(* IEC 61131-3 sources: llm-plc-st-eval/data/processed_definitivo/gemini-3.1-pro-preview/I5/zero_shot, 3 files *)

(* ---- ejec_1.st ---- *)
FUNCTION_BLOCK FB_Clasificadora
VAR_INPUT
    sensorPresencia : BOOL; // Sensor que detecta el paso de una pieza
    sensorAltura : BOOL;    // Sensor que detecta si la pieza es alta
END_VAR

VAR_OUTPUT
    banda : BOOL;           // Salida para activar la banda transportadora
    piston : BOOL;          // Salida para activar el pistón desviador
    nAltas : INT := 0;      // Contador de piezas altas
    nBajas : INT := 0;      // Contador de piezas bajas
END_VAR

VAR
    trigPresencia : R_TRIG; // Detector de flanco de subida para el sensor de presencia
    esperaPiston : BOOL;    // Marca de memoria para iniciar el retardo del pistón
    tonRetardo : TON;       // Temporizador de retardo (llegada al desviador)
    tpPiston : TP;          // Temporizador de pulso (duración de activación del pistón)
END_VAR

// 1. La banda funciona continuamente
banda := TRUE;

// 2. Detección del paso de una pieza (flanco de subida)
trigPresencia(CLK := sensorPresencia);

IF trigPresencia.Q THEN
    IF sensorAltura THEN
        // Es una pieza alta
        nAltas := nAltas + 1;
        esperaPiston := TRUE; // Se activa la bandera para iniciar el retardo
    ELSE
        // Es una pieza baja
        nBajas := nBajas + 1;
    END_IF;
END_IF;

// 3. Temporizador de retardo: espera 2 segundos a que la pieza llegue al pistón
tonRetardo(IN := esperaPiston, PT := T#2S);

// Al cumplirse los 2 segundos, se apaga la marca de espera
IF tonRetardo.Q THEN
    esperaPiston := FALSE;
END_IF;

// 4. Temporizador de pulso: activa el pistón durante 1 segundo
// Se dispara con el flanco de subida de tonRetardo.Q
tpPiston(IN := tonRetardo.Q, PT := T#1S);

// 5. Asignación de la salida física del pistón
piston := tpPiston.Q;

END_FUNCTION_BLOCK

(* ---- ejec_2.st ---- *)
FUNCTION_BLOCK FB_Clasificadora
VAR_INPUT
    sensorPresencia : BOOL; (* Detecta el paso de una pieza *)
    sensorAltura    : BOOL; (* Detecta si la pieza es alta *)
END_VAR
VAR_OUTPUT
    banda   : BOOL; (* Control de la banda transportadora *)
    piston  : BOOL; (* Control del pistón desviador *)
    nAltas  : INT;  (* Contador de piezas altas *)
    nBajas  : INT;  (* Contador de piezas bajas *)
END_VAR
VAR
    flancoPresencia : R_TRIG; (* Detector de flanco para contar solo una vez por pieza *)
    esperaPiston    : BOOL;   (* Marca para iniciar el retardo del pistón *)
    timerRetardo    : TON;    (* Temporizador para el tiempo de viaje (2s) *)
    timerPiston     : TP;     (* Temporizador para la duración del pistón (1s) *)
END_VAR

(* La banda está siempre activa *)
banda := TRUE;

(* Detectar el flanco de subida del sensor de presencia *)
flancoPresencia(CLK := sensorPresencia);

(* Lógica de clasificación y conteo al detectar una pieza *)
IF flancoPresencia.Q THEN
    IF sensorAltura THEN
        nAltas := nAltas + 1;
        esperaPiston := TRUE; (* Activa la bandera para iniciar el retardo *)
    ELSE
        nBajas := nBajas + 1;
    END_IF;
END_IF;

(* Temporizador TON: espera 2 segundos desde que se detecta la pieza alta *)
timerRetardo(IN := esperaPiston, PT := T#2S);

(* Cuando pasan los 2 segundos, se resetea la marca de espera *)
IF timerRetardo.Q THEN
    esperaPiston := FALSE;
END_IF;

(* Temporizador TP: genera un pulso de 1 segundo para el pistón *)
(* Se dispara exactamente cuando timerRetardo.Q se activa *)
timerPiston(IN := timerRetardo.Q, PT := T#1S);

(* Asignar la salida del temporizador al pistón *)
piston := timerPiston.Q;

END_FUNCTION_BLOCK

(* ---- ejec_3.st ---- *)
FUNCTION_BLOCK FB_Clasificadora
VAR_INPUT
    sensorPresencia : BOOL; (* Sensor que detecta el paso de una pieza *)
    sensorAltura : BOOL;    (* Sensor que detecta si la pieza es alta *)
END_VAR

VAR_OUTPUT
    banda : BOOL;           (* Salida para activar la banda transportadora *)
    piston : BOOL;          (* Salida para activar el pistón desviador *)
    nAltas : INT := 0;      (* Contador de piezas altas *)
    nBajas : INT := 0;      (* Contador de piezas bajas *)
END_VAR

VAR
    trigPresencia : R_TRIG; (* Detector de flanco de subida para la presencia *)
    tonRetardo : TON;       (* Temporizador para el retardo de 2 segundos *)
    tpPiston : TP;          (* Temporizador de pulso para el pistón de 1 segundo *)
    esperandoPiston : BOOL := FALSE; (* Memoria para el retardo del pistón *)
END_VAR

(* 1. La banda funciona continuamente *)
banda := TRUE;

(* 2. Detección de nueva pieza (flanco de subida) *)
trigPresencia(CLK := sensorPresencia);

IF trigPresencia.Q THEN
    IF sensorAltura THEN
        (* Es una pieza alta *)
        nAltas := nAltas + 1;
        esperandoPiston := TRUE; (* Inicia el proceso de desvío *)
    ELSE
        (* Es una pieza baja *)
        nBajas := nBajas + 1;
    END_IF;
END_IF;

(* 3. Temporizador de retardo (2 segundos hasta llegar al desviador) *)
tonRetardo(IN := esperandoPiston, PT := T#2S);

(* Al cumplirse el tiempo de retardo, reseteamos la memoria de espera *)
IF tonRetardo.Q THEN
    esperandoPiston := FALSE;
END_IF;

(* 4. Temporizador del pistón (pulso de 1 segundo) *)
(* Se dispara con el flanco de subida de tonRetardo.Q *)
tpPiston(IN := tonRetardo.Q, PT := T#1S);

(* 5. Activación de la salida del pistón *)
piston := tpPiston.Q;

END_FUNCTION_BLOCK
